// TIA Portal V21 export
// export: Created 2026-11-10T19:11:29.4474563Z, ExportSetting WithDefaults, DisplayName Totally Integrated Automation Portal, DisplayVersion V21 Update 3, DisplayName STEP 7 Professional, DisplayVersion V21 Update 3, DisplayName STEP 7 Safety, DisplayVersion V21, DisplayName Tech WebApplication, DisplayVersion V21, DisplayName WinCC Basic/Comfort/Advanced, DisplayVersion V21 Update 3, DisplayName WinCC Unified, DisplayVersion V21 Update 3
DATA_BLOCK "FB_SysMulti_DB"   // DB6
VERSION : 0.1
// stored: AutoNumber true, DBAccessibleFromOPCUA true, DBAccessibleFromWebserver true, InstanceOfName FB_SysMulti, InstanceOfType FB
"FB_SysMulti"
   // VAR
   //    mTON_TIME { S7_SetPoint := 'True'} : TON_TIME;
   //    mTOF_TIME { S7_SetPoint := 'True'} : TOF_TIME;
   //    mTP_TIME { S7_SetPoint := 'True'} : TP_TIME;
   //    mTONR_TIME { S7_SetPoint := 'True'} : TONR_TIME;
   //    mTON_LTIME { S7_SetPoint := 'True'} : TON_LTIME;
   //    mTOF_LTIME { S7_SetPoint := 'True'} : TOF_LTIME;
   //    mTP_LTIME { S7_SetPoint := 'True'} : TP_LTIME;
   //    mTONR_LTIME { S7_SetPoint := 'True'} : TONR_LTIME;
   //    mCTU_INT { S7_SetPoint := 'True'} : CTU_INT;
   //    mCTD_INT { S7_SetPoint := 'True'} : CTD_INT;
   //    mCTUD_INT { S7_SetPoint := 'True'} : CTUD_INT;
   //    mCTU_SINT { S7_SetPoint := 'True'} : CTU_SINT;
   //    mCTU_DINT { S7_SetPoint := 'True'} : CTU_DINT;
   //    mCTU_LINT { S7_SetPoint := 'True'} : CTU_LINT;
   //    mCTU_UINT { S7_SetPoint := 'True'} : CTU_UINT;
   //    mCTU_USINT { S7_SetPoint := 'True'} : CTU_USINT;
   //    mCTU_UDINT { S7_SetPoint := 'True'} : CTU_UDINT;
   //    mCTU_ULINT { S7_SetPoint := 'True'} : CTU_ULINT;
   //    mCTD_DINT { S7_SetPoint := 'True'} : CTD_DINT;
   //    mCTUD_DINT { S7_SetPoint := 'True'} : CTUD_DINT;
   //    mCTUD_LINT { S7_SetPoint := 'True'} : CTUD_LINT;
   //    mCTUD_UDINT { S7_SetPoint := 'True'} : CTUD_UDINT;
   //    mR_TRIG { S7_SetPoint := 'True'} : R_TRIG;
   //    mF_TRIG { S7_SetPoint := 'True'} : F_TRIG;
   //    mTSEND_C { S7_SetPoint := 'True'} : TSEND_C;
   //    mTRCV_C { S7_SetPoint := 'True'} : TRCV_C;
   //    mTCON { S7_SetPoint := 'True'} : TCON;
   //    mTDISCON { S7_SetPoint := 'True'} : TDISCON;
   //    mTSEND { S7_SetPoint := 'True'} : TSEND;
   //    mTRCV { S7_SetPoint := 'True'} : TRCV;
   //    mTUSEND { S7_SetPoint := 'True'} : TUSEND;
   //    mTURCV { S7_SetPoint := 'True'} : TURCV;
   //    mTMAIL_C { S7_SetPoint := 'True'} : TMAIL_C;
   //    mT_CONFIG { S7_SetPoint := 'True'} : T_CONFIG;
   //    mGET { S7_SetPoint := 'True'} : GET;
   //    mPUT { S7_SetPoint := 'True'} : PUT;
   //    mUSEND { S7_SetPoint := 'True'} : USEND;
   //    mURCV { S7_SetPoint := 'True'} : URCV;
   //    mBSEND { S7_SetPoint := 'True'} : BSEND;
   //    mBRCV { S7_SetPoint := 'True'} : BRCV;
   //    mMB_CLIENT { S7_SetPoint := 'True'} : MB_CLIENT;
   //    mMB_SERVER { S7_SetPoint := 'True'} : MB_SERVER;
   //    mRDREC { S7_SetPoint := 'True'} : RDREC;
   //    mWRREC { S7_SetPoint := 'True'} : WRREC;
   //    mRALRM { S7_SetPoint := 'True'} : RALRM;
   //    mGETIO { S7_SetPoint := 'True'} : GETIO;
   //    mSETIO { S7_SetPoint := 'True'} : SETIO;
   //    mGETIO_PART { S7_SetPoint := 'True'} : GETIO_PART;
   //    mSETIO_PART { S7_SetPoint := 'True'} : SETIO_PART;
   //    mProgram_Alarm { S7_SetPoint := 'True'} : Program_Alarm;
   //    mDRUM { S7_SetPoint := 'True'} : DRUM;
   //    mDCAT { S7_SetPoint := 'True'} : DCAT;
   //    mMCAT { S7_SetPoint := 'True'} : MCAT;
   //    mIMC { S7_SetPoint := 'True'} : IMC;
   //    mSMC { S7_SetPoint := 'True'} : SMC;
   //    mLEAD_LAG { S7_SetPoint := 'True'} : LEAD_LAG;
   //    mPID_Compact { S7_SetPoint := 'True'} : PID_Compact;
   //    mPID_3Step { S7_SetPoint := 'True'} : PID_3Step;
   //    mPID_Temp { S7_SetPoint := 'True'} : PID_Temp;
   //    mCONT_C { S7_SetPoint := 'True'} : CONT_C;
   //    mCONT_S { S7_SetPoint := 'True'} : CONT_S;
   //    mPULSEGEN { S7_SetPoint := 'True'} : PULSEGEN;
   //    mTCONT_CP { S7_SetPoint := 'True'} : TCONT_CP;
   //    mTCONT_S { S7_SetPoint := 'True'} : TCONT_S;
   //    aTon { S7_SetPoint := 'True'} : Array[0..1] of TON_TIME;
   //    aSend { S7_SetPoint := 'True'} : Array[0..1] of TSEND_C;
   // END_VAR
BEGIN
END_DATA_BLOCK
